(* IEC 61131-3 sources: codesys/project-view/Device/Plc Logic/Application/000-模组/向量阵列, 6 files *)

(* ---- IVectorArray.st ---- *)
INTERFACE IVectorArray
END_INTERFACE

//三点示教设置阵列参数
METHOD METH_SetPara : BOOL
VAR_INPUT
	Vector_O						: SMC_VECTOR3D;//工位原点坐标
	Vector_X						: SMC_VECTOR3D;//工位X轴终点坐标
	Vector_Y						: SMC_VECTOR3D;//工位Y轴终点坐标

	uiColumn_X						: UINT;//X轴方向工位数/列数
	uiRow_Y							: UINT;//Y轴方向工位数/行数
END_VAR
END_METHOD

//直接输入单位向量设置阵列参数
//常用于单点示教阵列
METHOD METH_SetParaByUnitVector : BOOL
VAR_INPUT
	Vector_O						: SMC_VECTOR3D;//工位原点坐标
	UnitVector_X					: SMC_VECTOR3D;//X轴方向的单位向量
	UnitVector_Y					: SMC_VECTOR3D;//Y轴方向的单位向量

	uiColumn_X						: UINT;//X轴方向工位数/列数
	uiRow_Y							: UINT;//Y轴方向工位数/行数
END_VAR
END_METHOD

//清除错误
METHOD METH_ClearError : BOOL
VAR_INPUT
END_VAR
END_METHOD

//通过行列坐标获取目标位置，坐标从(0,0)开始
METHOD METH_GetPosByCoordinate : SMC_VECTOR3D
VAR_INPUT
	uiColumn_X						: UINT;//X轴方向工位数/列数
	uiRow_Y							: UINT;//Y轴方向工位数/行数
END_VAR
END_METHOD

//可用的阵列总数
METHOD METH_Sum : UINT
VAR_INPUT
	uiColumn_X						: UINT;//X轴方向工位数/列数
	uiRow_Y							: UINT;//Y轴方向工位数/行数
END_VAR
END_METHOD

//对角线示教设置矩形阵列参数
//因只有对角线2个点，不能确定一个平行四边形，所以此函数默认阵列是矩形
METHOD METH_SetParaWithDiagonalRectangle: BOOL
VAR_INPUT
	Vector_O						: SMC_VECTOR3D;//工位原点坐标
	Vector_E						: SMC_VECTOR3D;//工位终点坐标/对角坐标

	uiColumn_X						: UINT;//X轴方向工位数/列数
	uiRow_Y							: UINT;//Y轴方向工位数/行数
END_VAR
END_METHOD

//通过大于0的序号获取目标位置
METHOD METH_GetPosByPoint : SMC_VECTOR3D
VAR_INPUT
	uiNum							: UINT;//整列序号
END_VAR
END_METHOD

(* ---- FC_CoordinateToPoint.st ---- *)
//输入从(0,0)开始的坐标，返回从X轴数过去且从1开始的序号。
//输入设定的行数与列数均大于0；
//函数返回值>0，计算无误；返回值=0，输入数据错误。
FUNCTION FC_CoordinateToPoint : UINT
VAR_INPUT
	uiCoordinate_X					: UINT;//X轴坐标
	uiCoordinate_Y					: UINT;//Y轴坐标
	uiColumn_X						: UINT;//X轴方向工位数/列数
	uiRow_Y							: UINT;//Y轴方向工位数/行数
END_VAR

VAR
	i								: UINT;

END_VAR
// --- implementation ---
IF uiColumn_X=0 OR uiRow_Y=0 OR uiCoordinate_X>=uiColumn_X OR uiCoordinate_Y>=uiRow_Y THEN
	FC_CoordinateToPoint := 0;
	RETURN;
END_IF

IF uiColumn_X = 1 THEN	//只有从Y轴方向延伸的一列
	FC_CoordinateToPoint := uiCoordinate_Y + 1;

ELSE	//只有从X轴方向延伸的一行，或者是有行有列
	i := uiCoordinate_Y * uiColumn_X;					//算出已填满的行有多少个
	i := i + uiCoordinate_X;							//再算出未填满的那一行，有多少个
	FC_CoordinateToPoint := i + 1;						//因为输出的序号要从1开始，加补偿

END_IF
END_FUNCTION

(* ---- FC_PointToCoordinate.st ---- *)
//输入大于0的序号和行列数，根据行列数转换为第一象限坐标，坐标从(0,0)开始。
//函数返回true表示计算无误；
//函数返回false表示输入数据错误，输出坐标固定为(0,0)。
FUNCTION FC_PointToCoordinate : BOOL
VAR_INPUT
	uiTargetPoint					: UINT;//目标序号
	uiColumn_X						: UINT;//X轴方向工位数/列数
	uiRow_Y							: UINT;//Y轴方向工位数/行数
END_VAR

VAR_OUTPUT
	Coordinate_X					: UINT;//X轴坐标
	Coordinate_Y					: UINT;//Y轴坐标
END_VAR

VAR
	i								: UINT;
	Rounding						: UINT;//整数部分
	Remainder						: UINT;//余数
	tmpCoordinate_X					: UINT;//X轴坐标
	tmpCoordinate_Y					: UINT;//Y轴坐标
END_VAR
// --- implementation ---
IF uiColumn_X=0 OR uiRow_Y=0 OR uiTargetPoint=0 OR uiTargetPoint>uiColumn_X*uiRow_Y THEN
	RETURN;
END_IF

(****	下面算法适用于坐标从(1,1)开始，后面要转化	****)
Rounding := uiTargetPoint / uiColumn_X;//行序号
Remainder := uiTargetPoint MOD uiColumn_X;//最终停留的所在列序号

(*转化成从(0,0)开始的坐标*)
IF Remainder > 0 THEN	//有余数，表示下一行还有计算
	tmpCoordinate_X := Remainder - 1;
	tmpCoordinate_Y := Rounding;//本来行数+1，但转化成从(0,0)开始的坐标，所以不需要

ELSE					//没有余数，表示停留在最后一行的最后一列
	tmpCoordinate_X := uiColumn_X - 1;
	tmpCoordinate_Y := Rounding - 1;

END_IF

(*输出结果*)
Coordinate_X := tmpCoordinate_X;
Coordinate_Y := tmpCoordinate_Y;

FC_PointToCoordinate := TRUE;
END_FUNCTION

(* ---- FB_VectorArray.st ---- *)
//三维向量阵列
FUNCTION_BLOCK FB_VectorArray IMPLEMENTS IVectorArray
VAR_INPUT
END_VAR

VAR_OUTPUT
	uiSum							: UINT;//可用的阵列总数
	bHasInitPara					: BOOL;//标志位，已设置阵列参数
	iErrorCode						: INT;//错误码
END_VAR

VAR
	//点位
	Vector_O						: SMC_VECTOR3D;//工位原点坐标
	Vector_X						: SMC_VECTOR3D;//工位X轴终点坐标
	Vector_Y						: SMC_VECTOR3D;//工位Y轴终点坐标

	//行列数
	uiColumn_X						: UINT;//X轴方向工位数/列数
	uiRow_Y							: UINT;//Y轴方向工位数/行数

	//单位向量
	UnitVector_X					: SMC_VECTOR3D;//X轴方向的单位向量
	UnitVector_Y					: SMC_VECTOR3D;//Y轴方向的单位向量

	Vector_Null						: SMC_VECTOR3D;//空向量

END_VAR
// --- implementation ---
(*第一次使用该FB块，先调用 METH_SetPara() 或 METH_SetParaByUnitVector() 设置内部参数*)

(**********************************************************************************************************
bHasInitPara -> TRUE
表示已设置好实例化该FB的参数。

若在此基础上，重新设置参数，即再次调用METH_SetPara的时候，参数设置错误，iErrorCode会报错为1。
但是原本的阵列参数保持原来参数，不会改变

iErrorCode:
0	->	无错误
1	->	行列参数设置错误
2	->	该阵列工位还没有行列参数设置
3	->	行列索引超出原本设置的参数
4	->	行列坐标是屏蔽位置

***********************************************************************************************************)
END_FUNCTION_BLOCK

(*清除错误*)
METHOD METH_ClearError : BOOL
// --- implementation ---
iErrorCode := 0;
END_METHOD

(*通过行列坐标获取目标位置，坐标从(0,0)开始*)
METHOD METH_GetPosByCoordinate : SMC_VECTOR3D
VAR_INPUT
	(*X轴方向工位数/列数 *)
	uiColumn_X						: UINT;
	(*Y轴方向工位数/行数 *)
	uiRow_Y							: UINT;
END_VAR

VAR
	tmpVector_X						: SMC_VECTOR3D;
	tmpVector_Y						: SMC_VECTOR3D;
	tmpVector_T						: SMC_VECTOR3D;
	tmpVector_Null					: SMC_VECTOR3D;

END_VAR
// --- implementation ---
iErrorCode := 0;

//没有设置阵列参数
IF NOT bHasInitPara THEN
	iErrorCode := 2;
	RETURN;
END_IF

//行列索引超出原本设置的参数
IF uiColumn_X > THIS^.uiColumn_X OR uiRow_Y > THIS^.uiRow_Y THEN
	iErrorCode := 3;
	RETURN;
END_IF

(****	根据行列点位，偏移单位向量，得出目标点位。从(0,0)开始	****)
IF uiColumn_X > 0 THEN
	//从原点偏移uiColumn_X个单位向量X
	SMC_V3_Mult(vDst:=tmpVector_X , vSrc:=UnitVector_X , d:=TO_LREAL(uiColumn_X) );
ELSE
	tmpVector_X := tmpVector_Null;
END_IF

IF uiRow_Y > 0 THEN
	//从原点偏移uiRow_Y个单位向量Y
	SMC_V3_Mult(vDst:=tmpVector_Y , vSrc:=UnitVector_Y , d:=TO_LREAL(uiRow_Y) );
ELSE
	tmpVector_Y := tmpVector_Null;
END_IF

SMC_V3_Add(vDst:=tmpVector_T , vLhs:=THIS^.Vector_O , vRhs:=tmpVector_X );
SMC_V3_Add(vDst:=tmpVector_T , vLhs:=tmpVector_T , vRhs:=tmpVector_Y );
METH_GetPosByCoordinate := tmpVector_T;
END_METHOD

(*通过大于0的序号获取目标位置*)
METHOD METH_GetPosByPoint : SMC_VECTOR3D
VAR_INPUT
	(*整列序号*)
	uiNum							: UINT;
END_VAR

VAR
	uiColumn_X						: UINT;
	uiRow_Y							: UINT;

	tmpVector_X						: SMC_VECTOR3D;
	tmpVector_Y						: SMC_VECTOR3D;
	tmpVector_T						: SMC_VECTOR3D;
	tmpVector_Null					: SMC_VECTOR3D;

	bFC_Done						: BOOL;
END_VAR
// --- implementation ---
iErrorCode := 0;

//没有设置阵列参数
IF NOT bHasInitPara THEN
	iErrorCode := 2;
	RETURN;
END_IF

//行列索引超出原本设置的参数
IF uiNum = 0 THEN
	iErrorCode := 3;
	RETURN;
END_IF

//序号转换成从(0,0)开始的坐标
bFC_Done := FC_PointToCoordinate(
				uiTargetPoint:=uiNum ,
				uiColumn_X:=THIS^.uiColumn_X ,
				uiRow_Y:=THIS^.uiRow_Y ,
				Coordinate_X=>uiColumn_X ,
				Coordinate_Y=>uiRow_Y );

IF NOT bFC_Done THEN//序号转换坐标失败，常见于uiNum值大于总阵列数
	iErrorCode := 3;
	RETURN;
END_IF

(****	根据行列点位，偏移单位向量，得出目标点位。从(0,0)开始	****)
IF uiColumn_X > 0 THEN
	//从原点偏移uiColumn_X个单位向量X
	SMC_V3_Mult(vDst:=tmpVector_X , vSrc:=UnitVector_X , d:=TO_LREAL(uiColumn_X) );
ELSE
	tmpVector_X := tmpVector_Null;
END_IF

IF uiRow_Y > 0 THEN
	//从原点偏移uiRow_Y个单位向量Y
	SMC_V3_Mult(vDst:=tmpVector_Y , vSrc:=UnitVector_Y , d:=TO_LREAL(uiRow_Y) );
ELSE
	tmpVector_Y := tmpVector_Null;
END_IF

SMC_V3_Add(vDst:=tmpVector_T , vLhs:=THIS^.Vector_O , vRhs:=tmpVector_X );
SMC_V3_Add(vDst:=tmpVector_T , vLhs:=tmpVector_T , vRhs:=tmpVector_Y );
METH_GetPosByPoint := tmpVector_T;
END_METHOD

(*三点示教设置阵列参数*)
METHOD METH_SetPara : BOOL
VAR_INPUT
	(*工位原点坐标*)
	Vector_O						: SMC_VECTOR3D;
	(*工位X轴终点坐标*)
	Vector_X						: SMC_VECTOR3D;
	(*工位Y轴终点坐标*)
	Vector_Y						: SMC_VECTOR3D;
	(*X轴方向工位数/列数 *)
	uiColumn_X						: UINT;
	(*Y轴方向工位数/行数 *)
	uiRow_Y							: UINT;
END_VAR

VAR
	//行列向量
	Vector_Xline					: SMC_VECTOR3D;
	Vector_Yline					: SMC_VECTOR3D;

END_VAR
// --- implementation ---
iErrorCode := 0;

(*行列数都是0，不是阵列，参数设置有误*)
IF uiColumn_X = 0 OR uiRow_Y = 0 THEN
	iErrorCode := 1;
	RETURN;
END_IF

(*向量相减，计算行列向量*)
SMC_V3_Sub(vDst:=Vector_Xline , vLhs:=Vector_X , vRhs:=Vector_O );
SMC_V3_Sub(vDst:=Vector_Yline , vLhs:=Vector_Y , vRhs:=Vector_O );

(****
根据行列数量，计算行列的单位向量
(uiColumn_X-1)和(uiRow_Y-1)都要减1，是因为这里算的是位置之间的间距数量，不是位置本身的数量
****)
IF uiColumn_X > 1 THEN
	SMC_V3_Mult(vDst:=UnitVector_X , vSrc:=Vector_Xline , d:=1 / TO_LREAL(uiColumn_X-1) );
ELSE
	UnitVector_X := Vector_Null;
END_IF

IF uiRow_Y > 1 THEN
	SMC_V3_Mult(vDst:=UnitVector_Y , vSrc:=Vector_Yline , d:=1 / TO_LREAL(uiRow_Y-1) );
ELSE
	UnitVector_Y := Vector_Null;
END_IF

(****	Meth形参赋值给FB实参	****)
THIS^.Vector_O := Vector_O;
THIS^.Vector_X := Vector_X;
THIS^.Vector_Y := Vector_Y;
THIS^.uiColumn_X := uiColumn_X;
THIS^.uiRow_Y := uiRow_Y;
uiSum := METH_Sum(uiColumn_X:=uiColumn_X , uiRow_Y:=uiRow_Y );//计算可用的阵列总数
bHasInitPara := TRUE;//标志位置true，已设置该FB阵列参数

METH_SetPara := TRUE;
END_METHOD

(*直接输入单位向量设置阵列参数
常用于单点示教阵列*)
METHOD METH_SetParaByUnitVector : BOOL
VAR_INPUT
	(*工位原点坐标*)
	Vector_O						: SMC_VECTOR3D;
	(*X轴方向的单位向量*)
	UnitVector_X					: SMC_VECTOR3D;
	(*Y轴方向的单位向量*)
	UnitVector_Y					: SMC_VECTOR3D;
	(*X轴方向工位数/列数 *)
	uiColumn_X						: UINT;
	(*Y轴方向工位数/行数 *)
	uiRow_Y							: UINT;
END_VAR

VAR
	//行列向量
	Vector_Xline					: SMC_VECTOR3D;
	Vector_Yline					: SMC_VECTOR3D;
END_VAR
// --- implementation ---
iErrorCode := 0;

(*行列数都是0，不是阵列，参数设置有误*)
IF uiColumn_X = 0 OR uiRow_Y = 0 THEN
	iErrorCode := 1;
	RETURN;
END_IF

(****	Meth形参赋值给FB实参	****)
THIS^.Vector_O := Vector_O;
THIS^.UnitVector_X := UnitVector_X;
THIS^.UnitVector_Y := UnitVector_Y;
THIS^.uiColumn_X := uiColumn_X;
THIS^.uiRow_Y := uiRow_Y;
uiSum := METH_Sum(uiColumn_X:=uiColumn_X , uiRow_Y:=uiRow_Y );//计算可用的阵列总数
bHasInitPara := TRUE;//标志位置true，已设置该FB阵列参数

METH_SetParaByUnitVector := TRUE;
END_METHOD

(*对角线示教设置阵列参数*)
(*因只有对角线2个点，不能确定一个平行四边形，所以此函数默认阵列是矩形*)
METHOD METH_SetParaWithDiagonalRectangle: BOOL
VAR_INPUT
	Vector_O						: SMC_VECTOR3D;//工位原点坐标
	Vector_E						: SMC_VECTOR3D;//工位终点坐标/对角坐标（dZ不处理）

	uiColumn_X						: UINT;//X轴方向工位数/列数
	uiRow_Y							: UINT;//Y轴方向工位数/行数
END_VAR

VAR
	//行列向量
	Vector_Xline					: SMC_VECTOR3D;
	Vector_Yline					: SMC_VECTOR3D;

	//行列终点向量
	Vector_Xend						: SMC_VECTOR3D;
	Vector_Yend						: SMC_VECTOR3D;

	//待确认：两点只能决定线而不能决定一个平面，因此dZ统一取Vector_O.dZ*)
END_VAR
// --- implementation ---
iErrorCode := 0;

(*行列数都是0，不是阵列，参数设置有误*)
IF uiColumn_X = 0 OR uiRow_Y = 0 THEN
	iErrorCode := 1;
	RETURN;
END_IF

(*利用对角线计算行与列的终点向量*)
// Vector_Xend := Vector_O;
// Vector_Yend := Vector_O;
//
// Vector_Xend.dX := Vector_E.dX;
// Vector_Yend.dY := Vector_E.dY;

Vector_Xend := Vector_E;
Vector_Xend.dY := Vector_O.dY;

Vector_Yend := Vector_E;
Vector_Yend.dX := Vector_O.dX;

(*向量相减，计算行列向量*)
SMC_V3_Sub(vDst:=Vector_Xline , vLhs:=Vector_Xend , vRhs:=Vector_O );
SMC_V3_Sub(vDst:=Vector_Yline , vLhs:=Vector_Yend , vRhs:=Vector_O );

(****
根据行列数量，计算行列的单位向量
(uiColumn_X-1)和(uiRow_Y-1)都要减1，是因为这里算的是位置之间的间距数量，不是位置本身的数量
****)
IF uiColumn_X > 1 THEN
	SMC_V3_Mult(vDst:=UnitVector_X , vSrc:=Vector_Xline , d:=1 / TO_LREAL(uiColumn_X-1) );
ELSE
	UnitVector_X := Vector_Null;
END_IF

IF uiRow_Y > 1 THEN
	SMC_V3_Mult(vDst:=UnitVector_Y , vSrc:=Vector_Yline , d:=1 / TO_LREAL(uiRow_Y-1) );
ELSE
	UnitVector_Y := Vector_Null;
END_IF

(****	Meth形参赋值给FB实参	****)
THIS^.Vector_O := Vector_O;
THIS^.Vector_X := Vector_X;
THIS^.Vector_Y := Vector_Y;
THIS^.uiColumn_X := uiColumn_X;
THIS^.uiRow_Y := uiRow_Y;
uiSum := METH_Sum(uiColumn_X:=uiColumn_X , uiRow_Y:=uiRow_Y );//计算可用的阵列总数
bHasInitPara := TRUE;//标志位置true，已设置该FB阵列参数

METH_SetParaWithDiagonalRectangle := TRUE;
END_METHOD

(*可用的阵列总数*)
METHOD METH_Sum : UINT
VAR_INPUT
	(*X轴方向工位数/列数 *)
	uiColumn_X							: UINT;
	(*Y轴方向工位数/行数 *)
	uiRow_Y								: UINT;
END_VAR
// --- implementation ---
IF uiColumn_X=1 AND uiRow_Y=1 THEN
	METH_Sum := 1;

ELSIF uiColumn_X>1 AND uiRow_Y=1 THEN//只有列数（即只有1行）
	METH_Sum := uiColumn_X;

ELSIF uiColumn_X=1 AND uiRow_Y>1 THEN//只有行数（即只有1列）
	METH_Sum := uiRow_Y;

ELSIF uiColumn_X>1 AND uiRow_Y>1 THEN
	METH_Sum := uiColumn_X * uiRow_Y;

END_IF
END_METHOD

(* ---- FB_VectorArrayWithShield.st ---- *)
{attribute 'enable_dynamic_creation'}
//三维向量阵列，编号可以屏蔽/跳过
FUNCTION_BLOCK FB_VectorArrayWithShield EXTENDS FB_VectorArray
VAR_IN_OUT
	auiShield							: ARRAY[0..19] OF UINT;//屏蔽编号
END_VAR

VAR_INPUT
END_VAR

VAR_OUTPUT
END_VAR

VAR
	uiShieldSum							: UINT;//被屏蔽的数量
	uiOriSum							: UINT;//此阵列的原始数量（含屏蔽）

END_VAR
// --- implementation ---
// //屏蔽数组没有外部变量传入引用
// IF auiShield = 0 THEN
// 	iErrorCode := 5;
// 	RETURN;
// END_IF
//
//
// diShield_Low := LOWER_BOUND(auiShield , 1);
// diShield_High := UPPER_BOUND(auiShield , 1);
// diShieldNum := ABS(diShield_High - diShield_Low);
//
//
// //第一次有效初始化 或 屏蔽数组发生改变
// IF NOT bFirstOn THEN
// 	bFirstOn := TRUE;
// END_IF

//auiShield_Sort := auiShield;
END_FUNCTION_BLOCK

(*通过大于0的序号获取目标位置*)
METHOD METH_GetPosByPoint : SMC_VECTOR3D
VAR_INPUT
	(*整列序号*)
	uiNum									: UINT;
END_VAR

VAR
	uiUsed									: DINT;//可使用的数量
	uiOffset								: UINT;//经过偏移的值（跳过屏蔽序号的实际序号）
	i										: UINT;

END_VAR
// --- implementation ---
//根据屏蔽编号计算偏移值
FOR i := 1 TO uiOriSum DO
	IF NOT METH_IsShield(i) THEN		//每次去屏蔽数组轮询，查看是否被屏蔽
		uiUsed := uiUsed + 1;			//该阵列无屏蔽，可以使用，则+1
		IF uiUsed = uiNum THEN			//uiUsed = uiNum，表示已到目标序号
			uiOffset := i;
			EXIT;
		END_IF

	END_IF
END_FOR

METH_GetPosByPoint := SUPER^.METH_GetPosByPoint(uiNum:= uiOffset);
END_METHOD

(*清除错误*)
METHOD METH_ClearError : BOOL
// --- implementation ---
SUPER^.METH_ClearError();
END_METHOD

(*通过行列坐标获取目标位置，坐标从(0,0)开始*)
METHOD METH_GetPosByCoordinate : SMC_VECTOR3D
VAR_INPUT
	(*X轴方向工位数/列数 *)
	uiColumn_X								: UINT;
	(*Y轴方向工位数/行数 *)
	uiRow_Y									: UINT;
END_VAR

VAR
	i										: DINT;
	uiNum									: UINT;

END_VAR
// --- implementation ---
//不考虑屏蔽位置，计算输入坐标在绝对阵列中的编号
uiNum := FC_CoordinateToPoint(
						uiCoordinate_X	:= uiColumn_X,
						uiCoordinate_Y	:= uiRow_Y,
						uiColumn_X		:= SUPER^.uiColumn_X,
						uiRow_Y			:= SUPER^.uiRow_Y);

//查询屏蔽数组，若屏蔽数组的元素值有uiNum的值，则表示输入坐标是一个屏蔽位，报错返回
FOR i := LOWER_BOUND(auiShield , 1) TO UPPER_BOUND(auiShield , 1) DO
	IF auiShield[i]<>0 AND auiShield[i]=uiNum THEN
		iErrorCode := 4;
		RETURN;
	END_IF

END_FOR

//使用绝对阵列中的编号，调用父类方法 METH_GetPosByPoint （用标号获取坐标）
METH_GetPosByCoordinate := SUPER^.METH_GetPosByPoint(uiNum:= uiNum);
END_METHOD

//是否被屏蔽
METHOD METH_IsShield : BOOL
VAR_INPUT
	uiNum							: UINT;
END_VAR

VAR
	i								: DINT;

END_VAR
// --- implementation ---
FOR i := LOWER_BOUND(auiShield , 1) TO UPPER_BOUND(auiShield , 1) DO
	IF uiNum = auiShield[i] THEN
		METH_IsShield := TRUE;
		RETURN;
	END_IF

END_FOR
END_METHOD

(*三点示教设置阵列参数*)
METHOD METH_SetPara : BOOL
VAR_INPUT
	(*工位原点坐标*)
	Vector_O	: SMC_VECTOR3D;
	(*工位X轴终点坐标*)
	Vector_X	: SMC_VECTOR3D;
	(*工位Y轴终点坐标*)
	Vector_Y	: SMC_VECTOR3D;
	(*X轴方向工位数/列数 *)
	uiColumn_X	: UINT;
	(*Y轴方向工位数/行数 *)
	uiRow_Y		: UINT;
END_VAR
// --- implementation ---
METH_SetPara := SUPER^.METH_SetPara(
							Vector_O		:= Vector_O	,
							Vector_X		:= Vector_X	,
							Vector_Y		:= Vector_Y	,
							uiColumn_X		:= uiColumn_X	,
							uiRow_Y			:= uiRow_Y		);

//auiShield_Sort := auiShield;
//OSCAT_BASIC._ARRAY_SORT(PT:=ADR(auiShield_Sort) , SIZE:=SIZEOF(auiShield_Sort) );
uiSum := METH_Sum(uiColumn_X:=uiColumn_X , uiRow_Y:=uiRow_Y );//计算可用的阵列总数
END_METHOD

(*直接输入单位向量设置阵列参数
常用于单点示教阵列*)
METHOD METH_SetParaByUnitVector : BOOL
VAR_INPUT
	(*工位原点坐标*)
	Vector_O		: SMC_VECTOR3D;
	(*X轴方向的单位向量*)
	UnitVector_X	: SMC_VECTOR3D;
	(*Y轴方向的单位向量*)
	UnitVector_Y	: SMC_VECTOR3D;
	(*X轴方向工位数/列数 *)
	uiColumn_X	: UINT;
	(*Y轴方向工位数/行数 *)
	uiRow_Y	: UINT;
END_VAR
// --- implementation ---
METH_SetParaByUnitVector := SUPER^.METH_SetParaByUnitVector(
													Vector_O		:= Vector_O	,
													UnitVector_X	:= UnitVector_X,
													UnitVector_Y	:= UnitVector_Y,
													uiColumn_X		:= uiColumn_X	,
													uiRow_Y			:= uiRow_Y		);

//auiShield_Sort := auiShield;
//OSCAT_BASIC._ARRAY_SORT(PT:=ADR(auiShield_Sort) , SIZE:=SIZEOF(auiShield_Sort) );
uiSum := METH_Sum(uiColumn_X:=uiColumn_X , uiRow_Y:=uiRow_Y );//计算可用的阵列总数
END_METHOD

(*对角线示教设置阵列参数*)
(*因只有对角线2个点，不能确定一个平行四边形，所以此函数默认阵列是矩形*)
METHOD METH_SetParaWithDiagonalRectangle: BOOL
VAR_INPUT
	Vector_O						: SMC_VECTOR3D;//工位原点坐标
	Vector_E						: SMC_VECTOR3D;//工位终点坐标/对角坐标（dZ不处理）

	uiColumn_X						: UINT;//X轴方向工位数/列数
	uiRow_Y							: UINT;//Y轴方向工位数/行数
END_VAR

VAR
	//行列向量
	Vector_Xline					: SMC_VECTOR3D;
	Vector_Yline					: SMC_VECTOR3D;

	//行列终点向量
	Vector_Xend						: SMC_VECTOR3D;
	Vector_Yend						: SMC_VECTOR3D;

END_VAR
// --- implementation ---
METH_SetParaWithDiagonalRectangle := SUPER^.METH_SetParaWithDiagonalRectangle(
												Vector_O	:= Vector_O	,
												Vector_E	:= Vector_E	,
												uiColumn_X	:= uiColumn_X	,
												uiRow_Y		:= uiRow_Y		);

//auiShield_Sort := auiShield;
//OSCAT_BASIC._ARRAY_SORT(PT:=ADR(auiShield_Sort) , SIZE:=SIZEOF(auiShield_Sort) );
uiSum := METH_Sum(uiColumn_X:=uiColumn_X , uiRow_Y:=uiRow_Y );//计算可用的阵列总数
END_METHOD

(*可用的阵列总数*)
METHOD METH_Sum : UINT
VAR_INPUT
	(*X轴方向工位数/列数 *)
	uiColumn_X							: UINT;
	(*Y轴方向工位数/行数 *)
	uiRow_Y								: UINT;
END_VAR

VAR
	i,j									: DINT;

END_VAR
// --- implementation ---
//先算出不带屏蔽的原始数量
uiOriSum := SUPER^.METH_Sum(uiColumn_X:=uiColumn_X , uiRow_Y:=uiRow_Y);

//计算被屏蔽的数量
uiShieldSum := 0;
FOR i := LOWER_BOUND(auiShield , 1) TO UPPER_BOUND(auiShield , 1) DO
	IF auiShield[i] <> 0 THEN
		uiShieldSum := uiShieldSum + 1;
	END_IF
END_FOR

//计算可用阵列的总数
uiSum := 0;
FOR i := 1 TO uiOriSum DO
	IF NOT METH_IsShield( TO_UINT(i) ) THEN
		uiSum := uiSum + 1;
	END_IF
END_FOR

METH_Sum := uiSum;
END_METHOD

(* ---- Example_VectorArray.st ---- *)
PROGRAM Example_VectorArray
VAR
	//向量阵列
	FB_50Array					: FB_VectorArray;					//50ml盘架
	FB_15Array					: FB_VectorArray;					//15ml盘架
	FB_15analArray				: FB_VectorArrayWithShield;			//15anal盘架

	auiShield					: ARRAY[0..19] OF UINT:=[4,6];//屏蔽编号，举例：4号和6号数学工位屏蔽

	//50ml试管盘架的单位向量（机械工位偏移）
	rRank50_X							: SMC_VECTOR3D:=(dX:=41,dY:=0,dZ:=0);
	rRank50_Y							: SMC_VECTOR3D:=(dX:=0,dY:=41,dZ:=0);

	//示教变量	[1..3]-->[原点坐标，X轴末端坐标，Y轴末端坐标]
	Pos_50								: ARRAY[1..3] OF SMC_VECTOR3D;//50ml示教试管管架位置
	Pos_15								: ARRAY[1..3] OF SMC_VECTOR3D;//15ml示教试管管架位置
	Pos_15anal							: ARRAY[1..3] OF SMC_VECTOR3D;//15ml示教分析试管管架位置

	bSetPosPara							: BOOL;//触发改写阵列数据

	bGetPosByNum						: BOOL;//获取位置触发--序号
	bGetPosByCoor						: BOOL;//获取位置触发--坐标
	uiNum								: UINT:=4;//序号
	GetPos_50							: SMC_VECTOR3D;//50ml目标试管管架位置
	GetPos_15							: SMC_VECTOR3D;//15ml目标试管管架位置
	GetPos_15anal						: SMC_VECTOR3D;//15ml目标分析试管管架位置

	bError								: BOOL;//FB阵列报错（如：获取参数有误）

END_VAR
// --- implementation ---
FB_50Array();
FB_15Array();
FB_15analArray(auiShield:= auiShield);

//设置阵列参数
IF bSetPosPara THEN
	bSetPosPara := FALSE;
	//uiColumn_X:= 6,uiRow_Y:= 10	意为6列10行，共60个工位

	//单点示教偏移
	FB_50Array.METH_SetParaByUnitVector(
		Vector_O:= Pos_50[1],
		UnitVector_X:= rRank50_X,
		UnitVector_Y:= rRank50_Y,
		uiColumn_X:= 6,
		uiRow_Y:= 10);

	//对角线示教，只能是矩形
	FB_15Array.METH_SetParaWithDiagonalRectangle(
		Vector_O:= Pos_15[1],
		Vector_E:= Pos_15[2],
		uiColumn_X:= 6,
		uiRow_Y:= 10);

	//三点示教
	FB_15analArray.METH_SetPara(
		Vector_O:= Pos_15anal[1],
		Vector_X:= Pos_15anal[2],
		Vector_Y:= Pos_15anal[3],
		uiColumn_X:= 6,
		uiRow_Y:= 10);

END_IF

//根据序号获取位置坐标
IF bGetPosByNum THEN
	bGetPosByNum := FALSE;

	GetPos_50 := FB_50Array.METH_GetPosByPoint(uiNum:= uiNum);
	GetPos_15 := FB_15Array.METH_GetPosByPoint(uiNum:= uiNum);

	//15anal的4号工位被屏蔽，所以返回5号工位坐标，即返回真正使用的工位坐标
	GetPos_15anal := FB_15analArray.METH_GetPosByPoint(uiNum:= uiNum);

END_IF

//根据坐标获取位置坐标，坐标从(0,0)开始
IF bGetPosByCoor THEN
	bGetPosByCoor := FALSE;

	//(uiColumn_X:=4 , uiRow_Y:=0)，意为第4列第1行

	GetPos_50 := FB_50Array.METH_GetPosByCoordinate(uiColumn_X:=4 , uiRow_Y:=0);
	GetPos_15 := FB_15Array.METH_GetPosByCoordinate(uiColumn_X:=4 , uiRow_Y:=0);

	//15anal的获取坐标是4号屏蔽位，会立刻报错
	GetPos_15anal := FB_15analArray.METH_GetPosByCoordinate(uiColumn_X:=3 , uiRow_Y:=0);

END_IF

//报错
bError := FB_50Array.iErrorCode<>0 OR FB_15Array.iErrorCode<>0 OR FB_15analArray.iErrorCode<>0;
END_PROGRAM
